Fanuc KAREL source: kb00164.KL

PROGRAM KB00164
%STACKSIZE=65535
%PRIORITY=65535
%NOLOCKGROUP
VAR
P1 : FILE
P2 : INTEGER
P3 : INTEGER
BEGIN
P2=1
P3=1
SET_FILE_POS(P1,P2,P3)
END KB00164
